# EPICS substitutions: adsApp/Db/FB_DriveVirtual.substitutions
file "FB_DriveVirtual_v1_01.template"
{
pattern
{P,      PORT,      A, P, VP,     VI, VN   }
{ADSTEST:,  ADS_1,  "", "" , Main.M, 1, "" }
}
